FUNCTION_BLOCK CD_TEST
VAR_INPUT
  P : BOOL;
  LDI : BOOL;
END_VAR
VAR
  c : CTD;
END_VAR
BEGIN
  c(CD := P, LD := LDI, PV := 2);
  //#ASSERT NOT (LDI AND c.Q) : Pok
END_FUNCTION_BLOCK
